(* IEC 61131-3 sources: codesys-framework/txt/application/WeVe Core (library)/50 Component, 1 file *)

(* ---- FB_Component.pou.st ---- *)
FUNCTION_BLOCK ABSTRACT FB_Component IMPLEMENTS I_Component
VAR_INPUT
END_VAR
VAR_OUTPUT
END_VAR
VAR
	_xBusy 		: BOOL;
	_xDone 		: BOOL;
	_sName 		: STRING := 'Undefined name';
	_scError 	: SC_Error;
END_VAR

// --- BEGIN IMPLEMENTATION ---
